Fanuc KAREL source: NC0041.KL

PROGRAM NC0041
%NOLOCKGROUP
ROUTINE R
VAR
  X : INTEGER
BEGIN
  X = 1
  SELECT X OF
    CASE(1):
      X = X + 2
    CASE(2):
      X = X + 3
    ELSE:
      SELECT X OF
        CASE(1):
          X = X + 2
        CASE(2):
          X = X + 3
        ELSE:
          SELECT X OF
            CASE(1):
              X = X + 2
            CASE(2):
              X = X + 3
            ELSE:
              SELECT X OF
                CASE(1):
                  X = X + 2
                CASE(2):
                  X = X + 3
                ELSE:
                  SELECT X OF
                    CASE(1):
                      X = X + 2
                    CASE(2):
                      X = X + 3
                    ELSE:
                      SELECT X OF
                        CASE(1):
                          X = X + 2
                        CASE(2):
                          X = X + 3
                        ELSE:
                          SELECT X OF
                            CASE(1):
                              X = X + 2
                            CASE(2):
                              X = X + 3
                            ELSE:
                              SELECT X OF
                                CASE(1):
                                  X = X + 2
                                CASE(2):
                                  X = X + 3
                                ELSE:
                                  SELECT X OF
                                    CASE(1):
                                      X = X + 2
                                    CASE(2):
                                      X = X + 3
                                    ELSE:
                                      SELECT X OF
                                        CASE(1):
                                          X = X + 2
                                        CASE(2):
                                          X = X + 3
                                        ELSE:
                                          SELECT X OF
                                            CASE(1):
                                              X = X + 2
                                            CASE(2):
                                              X = X + 3
                                            ELSE:
                                              SELECT X OF
                                                CASE(1):
                                                  X = X + 2
                                                CASE(2):
                                                  X = X + 3
                                                ELSE:
                                                  SELECT X OF
                                                    CASE(1):
                                                      X = X + 2
                                                    CASE(2):
                                                      X = X + 3
                                                    ELSE:
                                                      SELECT X OF
                                                        CASE(1):
                                                          X = X + 2
                                                        CASE(2):
                                                          X = X + 3
                                                        ELSE:
                                                          SELECT X OF
                                                            CASE(1):
                                                              X = X + 2
                                                            CASE(2):
                                                              X = X + 3
                                                            ELSE:
                                                              SELECT X OF
                                                                CASE(1):
                                                                  X = X + 2
                                                                CASE(2):
                                                                  X = X + 3
                                                                ELSE:
                                                                  SELECT X OF
                                                                    CASE(1):
                                                                      X = X + 2
                                                                    CASE(2):
                                                                      X = X + 3
                                                                    ELSE:
                                                                      SELECT X OF
                                                                        CASE(1):
                                                                          X = X + 2
                                                                        CASE(2):
                                                                          X = X + 3
                                                                        ELSE:
                                                                          SELECT X OF
                                                                            CASE(1):
                                                                              X = X + 2
                                                                            CASE(2):
                                                                              X = X + 3
                                                                            ELSE:
                                                                              SELECT X OF
                                                                                CASE(1):
                                                                                  X = X + 2
                                                                                CASE(2):
                                                                                  X = X + 3
                                                                                ELSE:
                                                                                  X = X + 1
                                                                              ENDSELECT
                                                                          ENDSELECT
                                                                      ENDSELECT
                                                                  ENDSELECT
                                                              ENDSELECT
                                                          ENDSELECT
                                                      ENDSELECT
                                                  ENDSELECT
                                              ENDSELECT
                                          ENDSELECT
                                      ENDSELECT
                                  ENDSELECT
                              ENDSELECT
                          ENDSELECT
                      ENDSELECT
                  ENDSELECT
              ENDSELECT
          ENDSELECT
      ENDSELECT
  ENDSELECT
END R
BEGIN
  R
END NC0041
